(* Logix 5000 project; controller CIP_14485201 vendor 1 type 14 code 216 rev 38.11; software revision 38.01 *)

TASK MainTask (continuous, watchdog 500 ms) : MainProgram

MODULES
   Local : vendor 1 type 14 code 216 (5069 0, rev 38.11)
END_MODULES

PROGRAM MainProgram   (* main routine MainRoutine *)

ROUTINE MainRoutine   (* ladder *)
END_ROUTINE
END_PROGRAM
